GLOBALCONSTANTS FMI (* Failure Mode Identifiers (FMI) for DTCs, ISO 11783-12 / SAE J1939-73 *)
  (* Standard: 61499-1 *)
  (* Version 1.0, 2026-11-17, Franz Höpfinger *)
  PACKAGE isobus::pgn::diag;
  VAR_GLOBAL CONSTANT
    ABOVE_NORMAL_MOST_SEVERE : USINT := 0; (* Above normal range - most severe *)
    BELOW_NORMAL_MOST_SEVERE : USINT := 1; (* Below normal range - most severe *)
    DATA_ERRATIC : USINT := 2; (* Data erratic, intermittent or incorrect *)
    VOLTAGE_HIGH : USINT := 3; (* Voltage above normal, or shorted to high source *)
    VOLTAGE_LOW : USINT := 4; (* Voltage below normal, or shorted to low source *)
    CURRENT_LOW_OPEN_CIRCUIT : USINT := 5; (* Current below normal or open circuit *)
    CURRENT_HIGH_GROUNDED : USINT := 6; (* Current above normal or grounded circuit *)
    MECHANICAL_NOT_RESPONDING : USINT := 7; (* Mechanical system not responding *)
    ABNORMAL_FREQUENCY : USINT := 8; (* Abnormal frequency or pulse width *)
    ABNORMAL_UPDATE_RATE : USINT := 9; (* Abnormal update rate *)
    ABNORMAL_RATE_OF_CHANGE : USINT := 10; (* Abnormal rate of change *)
    ROOT_CAUSE_UNKNOWN : USINT := 11; (* Root cause not known *)
    BAD_DEVICE : USINT := 12; (* Bad intelligent device or component *)
    OUT_OF_CALIBRATION : USINT := 13; (* Out of calibration *)
    SPECIAL_INSTRUCTIONS : USINT := 14; (* Special instructions *)
    ABOVE_NORMAL_LEAST_SEVERE : USINT := 15; (* Above normal range - least severe *)
    ABOVE_NORMAL_MODERATELY_SEVERE : USINT := 16; (* Above normal range - moderately severe *)
    BELOW_NORMAL_LEAST_SEVERE : USINT := 17; (* Below normal range - least severe *)
    BELOW_NORMAL_MODERATELY_SEVERE : USINT := 18; (* Below normal range - moderately severe *)
    RECEIVED_NETWORK_DATA_ERROR : USINT := 19; (* Received network data in error *)
    CONDITION_EXISTS : USINT := 31; (* Condition exists *)
  END_VAR
END_GLOBALCONSTANTS
